TYPE Profiling_Station_DUT :
STRUCT
	Start:  BOOL;
	Ready:  BOOL;
	Running:  Bool;
	Done:  Bool;
	Valid:  Bool;
	OverWidth:  Bool;
	OverHeight:  Bool;
	OverLength:  Bool;
	Error_ID:  Word;
END_STRUCT
END_TYPE

(* stored: Version 1.1.0.1
   DUT Profiling_Station_DUT: Id {a0df741a-86eb-4f8f-b8dd-4115eb2ef365} *)
